(* IEC 61131-3 sources: sis-interlock-demo/tests/POUs/Helpers/FB_CemRig, 5 files *)

(* ---- FB_CemRig.decl.st ---- *)
// Назначение: стенд тестов FB_CauseEffect: подменное время (старт LTIME#1H), журнал событий и
//             исполнитель матрицы; тест пишет входы, команды и конфигурацию стенда и вызывает
//             Cycle/Step/Run/PressReset.
// Автор:      kr0nsch
// Версия:     0.1.0
// Документ:   docs/DESIGN.md, раздел «12.3 Граничные случаи (вручную, команда A)»
// ВНИМАНИЕ:   код демонстрационный и не предназначен для систем безопасности. Реальная ПАЗ
//             требует определения SIL, сертифицированных аппаратных и программных средств
//             и валидации по ГОСТ Р МЭК 61511.
FUNCTION_BLOCK FB_CemRig
VAR_INPUT
    stCfg           : ST_CemCfg;        // конфигурация матрицы
    stCmd           : ST_CemCmd;        // команды HMI (ФБ сбрасывает)
    axCauseIn       : ARRAY[1..GVL_Const.SIS_CAUSES_MAX] OF BOOL;   // требования причин
    xOverridePermit : BOOL := TRUE;     // ключ разрешения обходов
    xResetHw        : BOOL;             // кнопка «Сброс ПАЗ»
END_VAR
VAR
    fbTime : PL.FB_FakeTime;            // подменное время
    fbLog  : FB_SisTestLog;             // журнал событий
    fbCem  : FB_CauseEffect;            // ФБ под тестом
END_VAR

(* ---- Out.method.decl.st ---- *)
// Выход следствия j: TRUE — под напряжением
METHOD Out : BOOL
VAR_INPUT
    uiEffect : UINT;   // индекс следствия
END_VAR

(* ---- Run.method.decl.st ---- *)
// Шаги tStep до tDuration (последний — остаток), вызов после каждого шага; не больше 1500 шагов
METHOD Run
VAR_INPUT
    tDuration : TIME;   // сколько времени пройти
    tStep     : TIME;   // шаг
END_VAR
VAR
    tLeft  : TIME;      // осталось
    tNow   : TIME;      // этот шаг
    uiIter : UINT;      // шагов сделано
END_VAR

(* ---- SetNow.method.decl.st ---- *)
// Установить подменное время (в том числе назад)
METHOD SetNow
VAR_INPUT
    ltValue : LTIME;   // новое время
END_VAR

(* ---- Step.method.decl.st ---- *)
// Продвинуть время на шаг и вызвать FB_CauseEffect
METHOD Step
VAR_INPUT
    tStep : TIME;   // шаг времени
END_VAR
